(* IEC 61131-3 sources: daoli-st-library/DL_Process, 610 files *)

(* ---- FB_DL_AutoclaveSterilSeq.st ---- *)
(*==============================================================================
 * 组件名称 (Component)  : FB_DL_AutoclaveSterilSeq
 * 所属子库 (Sublibrary) : DL_Process
 * 当前版本 (Version)    : 1.0.1
 * 兼容性   (Platform)   : CODESYS 3.5+ / TwinCAT 3 / 汇川 InoProShop / 施耐德 Machine Expert
 *                         仅依赖 Standard.library（TON / R_TRIG / ABS），零厂商私有库
 * 功能描述 (Function)   : 灭菌釜脉动真空灭菌七态顺控（GMP F0 值合规）：
 *                           ePulse     脉动置换：重复「抽真空-进蒸汽」nPulseCnt 次
 *                                      （tPulse 半周期交替，回合完成计数）；
 *                           eHeatUp    升温：温压入带（fTempSetC±fTempTolC ∧
 *                                      fPrSetKpa±fPrTolKpa）→ eSteril，tHeatTo 超时
 *                                      分码 eNoPr（压不起）/ eNoTemp（温不到）；
 *                           eSteril    保压灭菌：tSteril 到时 ∧ F0 累计达标 ∧ 温压在带内
 *                                      才过相；F0 累计 fF0Acc += fF0Rate×fCycle/60，
 *                                      **带内才累加、带外冻结不倒扣**（保守侧）；
 *                                      带外持续 tBandTmo → eFault eSterilBand；
 *                           eExhaustDry 排气干燥 tExhaust 到时 → eDone。
 *                         bStop 任一相回 eIdle 不记故障；bStop 保留 F0 累计
 *                         （_fF0Acc 不清零，同批次再启动接续累计，仅 bReset
 *                         上升沿清 F0）；bReset 上升沿清全部锁存（R311）。
 * 接口     (Interface)  : 输入 bStart/bStop/bReset、fPrKpa 釜压（kPa）、fTempC 腔温（℃）、
 *                         fPrSetKpa/fTempSetC 灭菌设定、fPrTolKpa/fTempTolC 带半宽、
 *                         tSteril 保压时长、tPulse 脉动半周期、tHeatTo/tBandTmo/tExhaust
 *                         各相窗、nPulseCnt 置换次数、fF0Min F0 目标（min）、fF0Rate
 *                         F0 速率系数（min/min）、fCycle 扫描周期（s）；输出 ePhase 七态、
 *                         fF0AccMin F0 累计（min）、四相指示 BOOL 组、bDone、eCause、
 *                         bError。
 * 边界     (Boundary)   : ① **属主边界（写死）：本件只做灭菌时序编排与 F0 累计闸，不驱动
 *                         蒸汽阀/真空泵/排水阀**；执行器由 IO 映射层按相指示位驱动。
 *                         ② 七态 CASE + ELSE 兜底 eFault（R6）；段间 TON 各自专用
 *                         （tonPulse/tonHeatTo/tonSteril/tonBandTmo/tonExhaust，R228A
 *                         命名豁免式），段 0 无条件刷新，IN 由当前相与带内判据派生。
 *                         ③ eCause 分码：eNoPr（升不起压）/ eNoTemp（温不到）/ eSterilBand
 *                         （带外跌出）/ eCfgIllegal（组态非法）/ ePhaseBad（兜底），
 *                         归因唯一（R190）。
 *                         ④ 温压非有限 → eFault eCause=eNoTemp 分码（规格指定）。
 *                         ⑤ 组态闸：nPulseCnt=0、任一相时间 <= T#0S、设定值/带宽非正、
 *                         fF0Min<0、fF0Rate<0 → 锁存 eFault eCfgIllegal。
 *                         ⑥ F0 带外冻结：TON IN 派生式（带内才计时与累加），带外不倒扣
 *                         （头注释声明保守侧语义）。
 *                         ⑦ 温压带判定浮点全用 <= / >= 容差比较，禁 = 判等（R28）。
 *                         ⑧ 零全局耦合（无 GVL / VAR_EXTERNAL / 物理地址）。
 * 分工声明 (Scope)      : 温度带判定语义与 `FB_DL_ToleranceWindow` 同思想，本件自带实现
 *                         不引用（规格定为不内嵌引用，独立验收）。
 * 来源标签 (Source Tag) : T2-2 ◐（LBP 工艺分层只借灭菌工序分类事实，F0 累计口径为 GMP
 *                         公开定义，零文本复制）
 * 码表     (Codes)      : 本件不占用任何全局数字码位。出口为 ENUM 七态 + LREAL 累计 +
 *                         BOOL 组 + ENUM 成因；数字码位待主控收口阶段统一派号。
 * 红线自检 (Redline)    : R1 ✓ 零 GVL/VAR_EXTERNAL ｜ R2 ✓ 零 %I/%Q/%M ｜ R3 ✓ 纯 IEC 61131-3
 *                         R4 ✓ 非有限分码 + 带内累加闸 + 组态闸 + 周期缺省闸 ｜ R5 ✓ 声明逐行同行双语注释
 *                         R6 ✓ 七态 CASE 含 ELSE ｜ R7 ✓ 五 TON/两 R_TRIG 段 0 无条件刷新
 * 修订历史 (Revision)   : 2026-11-20  v1.0.1  R50 返修 R2：头注释补声明
 *                         「bStop 保留 F0 累计」口径——bStop 中止只清脉动
 *                         计数与子态，_fF0Acc 不清零（同批次再启动接续累计），
 *                         仅 bReset 上升沿清 F0 累计；逻辑零改动，契约不变。
 *                         2026-11-20  v1.0.0  R48 首版（批次 4 · 序号 18）
 *                         验收向量：脉动计满进升温；温压入带 + F0 达标 + tSteril 到 →
 *                         过相；带外跌出冻结计时；tBandTmo 超时故障；bStop 中止不记故障。
 *==============================================================================*)

TYPE E_DL_AcsPhase :
(
    eIdle      := 0,    // 待机 / Idle
    ePulse     := 10,   // 脉动置换相 / Pulsing vacuum-steam phase
    eHeatUp    := 20,   // 升温相 / Heat-up phase
    eSteril    := 30,   // 保压灭菌相 / Sterilization hold phase
    eExhaustDry:= 40,   // 排气干燥相 / Exhaust and dry phase
    eDone      := 50,   // 程序完成 / Sequence done
    eFault     := 90    // 故障（等复位）/ Fault, awaiting reset
);
END_TYPE

TYPE E_DL_AcsCause :
(
    eNone       := 0,   // 无异常 / No anomaly
    eNoPr       := 1,   // 升不起压（升温相压力超时）/ Pressure fail in heat-up
    eNoTemp     := 2,   // 温不到 / 温压非有限（分码共用温度侧成因）/ Temperature fail or non-finite
    eSterilBand := 3,   // 灭菌带外跌出超时 / Sterilization band dropout timeout
    eCfgIllegal := 4,   // 组态非法 / Illegal configuration
    ePhaseBad   := 5    // 非法相位兜底 / Illegal phase fallback
);
END_TYPE

FUNCTION_BLOCK FB_DL_AutoclaveSterilSeq
VAR_INPUT
    bStart    : BOOL := FALSE;     // 启动沿（eIdle 入脉动相） [-] / Start edge
    bStop     : BOOL := FALSE;     // 中止（任一相回 eIdle，不记故障） [-] / Abort to idle, no fault
    bReset    : BOOL := FALSE;     // 复位，上升沿清全部锁存（R311） [-] / Reset, rising edge clears all latches
    fPrKpa    : LREAL := 0.0;      // 釜压实测 [kPa] / Chamber pressure [kPa]
    fTempC    : LREAL := 0.0;      // 腔温实测 [℃] / Chamber temperature [degC]
    fPrSetKpa : LREAL := 200.0;    // 灭菌压力设定，域 > 0 [kPa] / Sterilization pressure setpoint [kPa]
    fTempSetC : LREAL := 121.0;    // 灭菌温度设定，域 > 0 [℃] / Sterilization temperature setpoint [degC]
    fPrTolKpa : LREAL := 10.0;     // 压力带半宽，域 > 0 [kPa] / Pressure band half-width [kPa]
    fTempTolC : LREAL := 1.0;      // 温度带半宽，域 > 0 [℃] / Temperature band half-width [degC]
    tSteril   : TIME := T#30M;     // 保压灭菌时长，域 > T#0S [ms] / Sterilization hold duration [ms]
    tPulse    : TIME := T#2M;      // 脉动半周期（抽真空/进蒸汽各一段），域 > T#0S [ms] / Pulse half-period [ms]
    tHeatTo   : TIME := T#60M;     // 升温相超时，域 > T#0S [ms] / Heat-up timeout [ms]
    tBandTmo  : TIME := T#5M;      // 灭菌带外容忍窗，域 > T#0S [ms] / Band dropout tolerance [ms]
    tExhaust  : TIME := T#15M;     // 排气干燥时长，域 > T#0S [ms] / Exhaust-dry duration [ms]
    nPulseCnt : UDINT := 3;        // 脉动置换次数，域 >= 1（=0 组态闸） [次] / Pulse swap count
    fF0Min    : LREAL := 3.0;      // F0 灭菌值目标，域 >= 0 [min] / F0 target [min]
    fF0Rate   : LREAL := 1.0;      // F0 累计速率系数（带内每分钟 F0 增量），域 >= 0 [min/min] / F0 rate coefficient
    fCycle    : LREAL := 0.0;      // 扫描周期（<=0 用缺省） [s] / Scan cycle, default used when <= 0
END_VAR
VAR_OUTPUT
    ePhase    : E_DL_AcsPhase;     // 当前相出口 [-] / Present phase outlet
    fF0AccMin : LREAL;             // F0 累计输出（带内累加、带外冻结） [min] / F0 accumulated [min]
    bPulseActive   : BOOL;         // 脉动相指示 [-] / Pulse phase indicator
    bHeatUpActive  : BOOL;         // 升温相指示 [-] / Heat-up phase indicator
    bSterilActive  : BOOL;         // 灭菌相指示 [-] / Sterilization phase indicator
    bExhaustActive : BOOL;         // 排气干燥相指示 [-] / Exhaust phase indicator
    bDone     : BOOL;              // 程序完成（eDone 驻留指示） [-] / Sequence done indicator
    eCause    : E_DL_AcsCause;     // 成因出口（锁存回放，R189） / Cause outlet, latched
    bError    : BOOL;              // 故障标志 [-] / Error flag
END_VAR
VAR
    _eState    : E_DL_AcsPhase := E_DL_AcsPhase.eIdle;   // 内部相（CASE 唯一写入目标） / Internal phase
    _eCause    : E_DL_AcsCause := E_DL_AcsCause.eNone;   // 成因锁存量 / Latched cause
    _bFault    : BOOL;             // 故障锁存位（解除沿 = bReset 上升沿） / Latched fault bit
    _nPulseDone: UDINT := 0;       // 脉动回合完成计数 [次] / Completed pulse swaps
    _bPulseStm : BOOL;             // 脉动子态（FALSE=抽真空段 / TRUE=进蒸汽段） / Pulse sub-state
    _bInBand   : BOOL;             // 当拍温压带内判据 [-] / In-band this scan
    _bNonFin   : BOOL;             // 温压非有限当拍量 [-] / Non-finite measurands this scan
    _bCfgBad   : BOOL;             // 组态非法当拍量 [-] / Illegal configuration this scan
    _fCy       : LREAL;            // 当拍有效周期 [s] / Effective cycle this scan
    _fF0Acc    : LREAL := 0.0;     // F0 累计锁存 [min] / F0 accumulator latch
    _bBusyPrev : BOOL;             // 上拍运行快照（bDone 迁出用） / Busy snapshot
    tonPulse   : TON;              // 脉动半周期定时器，段 0 无条件调用 / Pulse half-period timer
    tonHeatTo  : TON;              // 升温超时定时器，段 0 无条件调用 / Heat-up timeout timer
    tonSteril  : TON;              // 保压灭菌计时定时器，段 0 无条件调用 / Sterilization hold timer
    tonBandTmo : TON;              // 带外容忍窗定时器，段 0 无条件调用 / Band dropout tolerance timer
    tonExhaust : TON;              // 排气干燥计时定时器，段 0 无条件调用 / Exhaust-dry timer
    rtStart    : R_TRIG;           // 启动沿实例，段 0 无条件调用 / Start edge instance
    rtReset    : R_TRIG;           // 复位沿实例，段 0 无条件调用 / Reset edge instance
END_VAR
VAR CONSTANT
    DL_ACS_CYDEF : LREAL := 0.01;    // 缺省扫描周期 [s] / Default scan cycle
    DL_ACS_SEC   : LREAL := 60.0;    // 分秒换算基 [s/min] / Second-per-minute base
    DL_ACS_ZERO  : LREAL := 0.0;     // 非有限差值判零基准 [-] / Non-finite difference zero base
    DL_ACS_UDMAX : UDINT := 4294967295;   // UDINT 上限（脉动计数饱和点） [次] / UDINT ceiling
END_VAR

(* —— 段 0：非有限判 + 组态闸 + 周期派生 + 五 TON 两沿无条件周期刷新 —— *)
_bNonFin := (fPrKpa <> fPrKpa) OR ((fPrKpa - fPrKpa) <> DL_ACS_ZERO)
         OR (fTempC <> fTempC) OR ((fTempC - fTempC) <> DL_ACS_ZERO);   // 温压非有限（R245） / Non-finite pressure and temperature
_bCfgBad := (nPulseCnt = 0) OR (fPrSetKpa <= 0.0) OR (fTempSetC <= 0.0)
         OR (fPrTolKpa <= 0.0) OR (fTempTolC <= 0.0)
         OR (tSteril <= T#0S) OR (tPulse <= T#0S) OR (tHeatTo <= T#0S)
         OR (tBandTmo <= T#0S) OR (tExhaust <= T#0S)
         OR (fF0Min < 0.0) OR (fF0Rate < 0.0);          // 组态域闸（含 nPulseCnt=0） / Configuration gate
IF fCycle > 0.0 THEN
    _fCy := fCycle;                                     // 组态周期有效 / Configured cycle valid
ELSE
    _fCy := DL_ACS_CYDEF;                               // 周期缺省兜底 / Default cycle fallback
END_IF
rtStart(CLK := bStart);                                 // 启动沿，每拍必调 / Start edge, every scan
rtReset(CLK := bReset);                                 // 复位沿，每拍必调 / Reset edge, every scan
tonPulse(IN := (_eState = E_DL_AcsPhase.ePulse) AND (NOT tonPulse.Q), PT := tPulse);   // 脉动半周期自复位窗（R188） / Pulse self-reset window
tonHeatTo(IN := (_eState = E_DL_AcsPhase.eHeatUp), PT := tHeatTo);   // 升温超时（进相计时，出相自复位） / Heat-up timeout
tonSteril(IN := (_eState = E_DL_AcsPhase.eSteril) AND _bInBand, PT := tSteril);   // 灭菌计时（带内才计时，带外冻结） / Sterilization timer, in-band gated
tonBandTmo(IN := (_eState = E_DL_AcsPhase.eSteril) AND (NOT _bInBand), PT := tBandTmo);   // 带外容忍窗 / Band dropout tolerance
tonExhaust(IN := (_eState = E_DL_AcsPhase.eExhaustDry), PT := tExhaust);   // 排气干燥计时 / Exhaust timer

(* —— 段 1：带内判据（非有限按带外处理并分码 eNoTemp，先于 CASE 使用） —— *)
_bInBand := (NOT _bNonFin)
         AND (ABS(fTempC - fTempSetC) <= fTempTolC)     // 温度带内（容差比较，禁 =） / Temperature in band
         AND (ABS(fPrKpa - fPrSetKpa) <= fPrTolKpa);    // 压力带内 / Pressure in band

(* —— 段 2：单拍量预清零（_eState/_eCause/_bFault/_n PulseDone/_fF0Acc 锁存量不入清单，R107） —— *)
bPulseActive := FALSE;                                  // 脉动相指示预清 / Pulse indicator preset
bHeatUpActive := FALSE;                                 // 升温相指示预清 / Heat-up indicator preset
bSterilActive := FALSE;                                 // 灭菌相指示预清 / Sterilization indicator preset
bExhaustActive := FALSE;                                // 排气相指示预清 / Exhaust indicator preset
bDone := FALSE;                                         // 完成指示预清 / Done preset
bError := FALSE;                                        // 故障标志预清（R45 配对） / Error flag preset

(* —— 段 3：组态闸入故障 —— *)
IF _bCfgBad AND (NOT _bFault) THEN
    _bFault := TRUE;                                    // 锁存 / Latch
    _eCause := E_DL_AcsCause.eCfgIllegal;               // 归因：组态非法 / Cause: illegal config
    _eState := E_DL_AcsPhase.eFault;                    // 入故障相 / Enter fault
END_IF

(* —— 段 4：迁出链（bStop 优先不记故障；bReset 清全部锁存 R311） —— *)
IF bStop AND (_eState <> E_DL_AcsPhase.eIdle) THEN
    IF _eState = E_DL_AcsPhase.eFault THEN
        _bFault := FALSE;                               // 停机优先：故障相允许被停机清出 / Stop wins over fault
        _eCause := E_DL_AcsCause.eNone;                 // 清成因 / Clear cause
    END_IF
    _nPulseDone := 0;                                   // 清脉动计数 / Clear pulse count
    _bPulseStm := FALSE;                                // 清脉动子态 / Clear pulse sub-state
    _eState := E_DL_AcsPhase.eIdle;                     // 回待机（不记故障） / Back to idle, no fault
END_IF
IF rtReset.Q THEN
    _bFault := FALSE;                                   // 清故障锁存（R311） / Clear fault latch
    _eCause := E_DL_AcsCause.eNone;                     // 清成因 / Clear cause
    _nPulseDone := 0;                                   // 清脉动计数 / Clear pulse count
    _bPulseStm := FALSE;                                // 清脉动子态 / Clear pulse sub-state
    _fF0Acc := 0.0;                                     // 清 F0 累计 / Clear F0 accumulator
    _eState := E_DL_AcsPhase.eIdle;                     // 回待机 / Back to idle
END_IF

(* —— 段 5：七态顺控（只在无故障时推进；温压非有限 → 故障分码 eNoTemp） —— *)
IF (NOT _bFault) AND (NOT _bCfgBad) AND (NOT bStop) THEN
    IF _bNonFin AND (_eState <> E_DL_AcsPhase.eIdle) AND (_eState <> E_DL_AcsPhase.eDone) THEN
        _bFault := TRUE;                                // 运行相温压非有限：故障锁存（规格④） / Non-finite in running phase: fault
        _eCause := E_DL_AcsCause.eNoTemp;               // 归因分码：温度侧 / Cause: temperature side
        _eState := E_DL_AcsPhase.eFault;                // 入故障相 / Enter fault
    ELSE
        CASE _eState OF

        E_DL_AcsPhase.eIdle:
            IF rtStart.Q THEN
                _nPulseDone := 0;                       // 启动清脉动计数 / Clear pulse count on start
                _bPulseStm := FALSE;                    // 启动回抽真空子段 / Start in vacuum sub-phase
                _eState := E_DL_AcsPhase.ePulse;        // 入脉动相 / Enter pulse phase
            END_IF

        E_DL_AcsPhase.ePulse:
            IF tonPulse.Q THEN
                _bPulseStm := NOT _bPulseStm;           // 半周期到：抽真空/进蒸汽交替 / Half period: toggle sub-phase
                IF NOT _bPulseStm THEN
                    IF _nPulseDone < DL_ACS_UDMAX THEN
                        _nPulseDone := _nPulseDone + 1; // 完成一个完整回合（真空→蒸汽→真空）计数 / Count full swap round
                    END_IF
                END_IF
                IF _nPulseDone >= nPulseCnt THEN
                    _eState := E_DL_AcsPhase.eHeatUp;   // 置换次数达标：进升温相 / Swaps done: enter heat-up
                END_IF
            END_IF

        E_DL_AcsPhase.eHeatUp:
            IF _bInBand THEN
                _eState := E_DL_AcsPhase.eSteril;       // 温压入带：进保压灭菌相 / In band: enter sterilization
            ELSIF tonHeatTo.Q THEN
                IF ABS(fPrKpa - fPrSetKpa) > fPrTolKpa THEN
                    _eCause := E_DL_AcsCause.eNoPr;     // 压力超带：升不起压 / Pressure out of band: no pressure
                ELSE
                    _eCause := E_DL_AcsCause.eNoTemp;   // 压力入带而温度不达：温不到 / Temperature short
                END_IF
                _bFault := TRUE;                        // 超时故障锁存 / Latch fault
                _eState := E_DL_AcsPhase.eFault;        // 入故障相 / Enter fault
            END_IF

        E_DL_AcsPhase.eSteril:
            IF _bInBand THEN
                _fF0Acc := _fF0Acc + fF0Rate * _fCy / DL_ACS_SEC;   // 带内 F0 累计（速率×周期/60） / In-band F0 accumulation
            END_IF
            (* 带外不倒扣不累加（保守侧，头注释⑥）；带外容忍窗由 tonBandTmo 监视 *)
            IF tonBandTmo.Q THEN
                _eCause := E_DL_AcsCause.eSterilBand;   // 带外跌出超时 / Band dropout timeout
                _bFault := TRUE;                        // 锁存 / Latch
                _eState := E_DL_AcsPhase.eFault;        // 入故障相 / Enter fault
            ELSIF tonSteril.Q AND (_fF0Acc >= fF0Min) AND _bInBand THEN
                _eState := E_DL_AcsPhase.eExhaustDry;   // 计时到 ∧ F0 达标 ∧ 带内：过相（禁浮点 =，>= 判据） / Pass criteria met
            END_IF

        E_DL_AcsPhase.eExhaustDry:
            IF tonExhaust.Q THEN
                _eState := E_DL_AcsPhase.eDone;         // 排气干燥到时：进完成相 / Exhaust done: enter done
            END_IF

        E_DL_AcsPhase.eDone:
            ;                                           // 完成相驻留：由 bReset / bStop 迁出 / Held, exits via reset or stop

        E_DL_AcsPhase.eFault:
            ;                                           // 故障相驻留：由迁出链处理 / Held by exit chain

        ELSE
            _eCause := E_DL_AcsCause.ePhaseBad;         // 非法相位兜底归因 / Illegal phase cause
            _bFault := TRUE;                            // 锁存 / Latch
            _eState := E_DL_AcsPhase.eFault;            // 强拉故障相 / Force fault

        END_CASE
    END_IF
END_IF

(* —— 段 6：完成脉冲（由"运行→eDone"沿派生，单拍，R34 两段式） —— *)
IF _bBusyPrev AND (_eState = E_DL_AcsPhase.eDone) THEN
    bDone := TRUE;                                      // 程序完成单拍指示 / Done pulse
END_IF
_bBusyPrev := (_eState <> E_DL_AcsPhase.eIdle)
          AND (_eState <> E_DL_AcsPhase.eDone)
          AND (_eState <> E_DL_AcsPhase.eFault);        // 运行中快照（本拍末） / Busy snapshot at body end

(* —— 段 7：出口单点映射（相指示与相别同源，R191） —— *)
bPulseActive   := (_eState = E_DL_AcsPhase.ePulse);     // 脉动相指示 / Pulse indicator
bHeatUpActive  := (_eState = E_DL_AcsPhase.eHeatUp);    // 升温相指示 / Heat-up indicator
bSterilActive  := (_eState = E_DL_AcsPhase.eSteril);    // 灭菌相指示 / Sterilization indicator
bExhaustActive := (_eState = E_DL_AcsPhase.eExhaustDry);   // 排气相指示 / Exhaust indicator
IF _eState = E_DL_AcsPhase.eDone THEN
    bDone := TRUE;                                      // 完成相驻留期保持指示（R191 名实双出口声明） / Done held while resident
END_IF
ePhase := _eState;                                      // 当前相出口 / Present phase outlet
fF0AccMin := _fF0Acc;                                   // F0 累计出口 / F0 outlet
eCause := _eCause;                                      // 成因出口 / Cause outlet
bError := _bFault OR _bCfgBad;                          // 故障标志 = 锁存或组态非法 / Error = latch or config

END_FUNCTION_BLOCK

(* ---- FB_DL_BatchDoseSeq.st ---- *)
(*
    FB_DL_BatchDoseSeq —— 批次定量给料顺控（预给/快给/慢给/落料/校验 五相）
    ------------------------------------------------------------------
    组件名称  : FB_DL_BatchDoseSeq
    分类      : DL_Process / Batching
    前缀      : FB_DL_
    版本      : 1.0.0
    溯源      : 借鉴点 —— ISA-88（ANSI/ISA-88.00.01）批次控制模型的
                「单元配方 / 相逻辑 / 相超时 / 批次判定」分层思想，以及定量给料
                行业通行的三段给料法（快给料逼近 + 慢给料精给 + 落料补偿）。
                本件只借鉴**相划分与判定顺序**这两项公开语义。
                clean-room 声明 —— 零代码行复制；状态机为本件自有 ENUM + CASE，
                定时仅用 IEC 61131-3 标准库 TON，沿检测仅用标准库 R_TRIG。
                许可证 —— 本件 MIT；来源标签 isa88 指标准术语与模型，
                标准文本不属代码，无许可继承关系。
    平台      : 纯 IEC 61131-3，CODESYS 3.5 / TwinCAT 3 / InoProShop / Machine Expert 通用
    作者      : 道莅代码库 · PLC编程专家（R70 构建轮 · 批 1 · N4）
    ------------------------------------------------------------------
    功能说明  : 单批次定量给料顺控。相序：
                eIdle 待机 → ePreDose 预给料（预给料阀开，到 fPreW 止）
                → eFastDose 快给料（快给料阀开，到 fFastW 止）
                → eSlowDose 慢给料（慢给料阀开，到 fTarget - fFreeFall 止）
                → eSettle 落料（全阀关，等 tSettle 让空中料落下）
                → eCheck 校验（净重对 fTarget ± 公差带判定）
                → eComplete 完成（保持，等下一次 bStart）。
                超时归因唯一（R190）：预给 / 快给 / 慢给 / 落料四相各持独立码
                0303 / 0304 / 0305 / 0306，绝不共用同一枚举或同一码值。
                定时器设计：单实例 _tonPhase，PT 由当前相在段 4 以 IF/ELSIF 链
                逐相选择（含 ELSE 缺省），**每周期无条件调用**（规则 ⑦），
                故选相不依赖任何可能被跳过的分支；落料相的正常出口也复用该
                实例的 Q（PT = tSettle），故落料相不存在「正常完成」与「超时」
                两种语义，只有「到时间进入校验」一种。
                相内比较全部用 >= 的闭区间口径，不用浮点相等（规则 ④）。
    错误码    : 16#0002_0301 组态非法（阈值不单调 / 负公差 / 非有限），清锁存后回 eIdle —— 故障级
                16#0002_0302 称重值非有限，锁存并停料 —— 故障级
                16#0002_0303 预给料相超时 —— 故障级
                16#0002_0304 快给料相超时 —— 故障级
                16#0002_0305 慢给料相超时 —— 故障级
                16#0002_0306 落料相超时 —— 故障级
                16#0002_0307 欠重（净重低于 fTarget - fTolNeg）—— 故障级
                16#0002_0308 超重（净重高于 fTarget + fTolPos）—— 故障级
                16#0002_0309 非法相枚举值（CASE ELSE 兜底）—— 故障级
                16#0002_0310 启动被拒（称斗未回零，fWeight 超过 fZeroTol）—— 信息级，不置 bError
    码位总账  : 0301 / 0302 / 0303 / 0304 / 0305 / 0306 / 0307 / 0308 / 0309 用（均故障级）
                0310 用（信息级，bError 恒 FALSE）
    状态机    : ENUM E_DL_BdsPhase 八态，CASE 全覆盖 + ELSE 兜底（回 eFault 并置 0309）。
                迁移表见功能说明；bAbort 任意相 → eIdle（操作态，不发码）；
                bReset 上升沿：解锁存 → eIdle（仅此一条可到达的解除边，R188）。
    边界与披露: 一 组态判据逐项点名（R272）：fTarget / fPreW / fFastW / fFreeFall /
                   fTolNeg / fTolPos 全部纳入非有限闸，并校验单调链
                   0 < fPreW < fFastW < (fTarget - fFreeFall) 与 fFreeFall < fTarget、
                   两侧公差 >= 0；任一不满足即 0301 并锁存，**不落任何阈值比较**；
                二 称重输入非有限即锁存 0302，全部给料出口立即关断（失效安全方向）；
                三 失能语义：本件无 bEn 引脚，停机由 bAbort 承担 —— bAbort 为电平
                   有效，任意拍为 TRUE 即回 eIdle 且输出全清零，不发码（操作态）；
                四 出口语义（R191 名实双出口）：bUnder / bOver 为校验相判定结果位，
                   同时映射到故障码 0307 / 0308 并锁存；eComplete 为完成相标志，
                   完成不算故障，bError 恒 FALSE；
                五 bBusy 定义：给料 / 落料 / 校验三区间（真正占用设备的时间窗）；
                   bValid 定义：出口可信（未处在锁存故障相）；
                六 定时器 _tonPhase 与沿实例 _rtStart / _rtReset 均无条件周期调用；
                七 零全局变量、零 VAR_EXTERNAL、零物理地址、零数组下标、无除法。
    修订记录  : 2026-11-22 v1.0.0 首次入库（R70 构建轮 · 批 1 · N4）
*)
TYPE E_DL_BdsPhase :
(
    eIdle     := 0,   (* 待机，等待启动 / idle, waiting for a start *)
    ePreDose  := 10,  (* 预给料相（大流量阀开）/ the pre-dose phase, the coarse valve open *)
    eFastDose := 20,  (* 快给料相（快给料阀开）/ the fast-dose phase, the fast valve open *)
    eSlowDose := 30,  (* 慢给料相（慢给料阀开）/ the slow-dose phase, the fine valve open *)
    eSettle   := 40,  (* 落料相（全阀关，等空中料落下）/ the settling phase, all valves closed *)
    eCheck    := 50,  (* 校验相（净重对公差带判定）/ the check phase, the net weight against the tolerance *)
    eComplete := 60,  (* 完成相（保持到下次启动）/ the complete phase, held until the next start *)
    eFault    := 70   (* 故障相（锁存待复位）/ the fault phase, latched for a reset *)
);
END_TYPE

FUNCTION_BLOCK FB_DL_BatchDoseSeq
VAR_INPUT
    bStart    : BOOL := FALSE;             (* 启动命令（上升沿有效），[标志] / the start command, rising edge effective *)
    bAbort    : BOOL := FALSE;             (* 中止命令（电平有效），[标志] / the abort command, level effective *)
    bReset    : BOOL := FALSE;             (* 故障复位（上升沿有效），[标志] / the fault reset, rising edge effective *)
    fWeight   : LREAL := 0.0;              (* 称斗净重实时值，[kg] / the live net weight of the weigh hopper *)
    fTarget   : LREAL := 25.0;             (* 批次目标净重，[kg]，须 > 0 / the batch target weight, must be positive *)
    fPreW     : LREAL := 5.0;              (* 预给料结束重量点，[kg]，须 < fFastW / the pre-dose hand-over weight *)
    fFastW    : LREAL := 20.0;             (* 快给料结束重量点，[kg]，须 < fTarget - fFreeFall / the fast-dose hand-over weight *)
    fFreeFall : LREAL := 1.0;              (* 慢给料提前关断量（空中落差），[kg]，须 < fTarget / the in-flight cut-off weight *)
    fTolNeg   : LREAL := 0.2;              (* 允许负偏差，[kg]，须 >= 0 / the permitted negative deviation *)
    fTolPos   : LREAL := 0.2;              (* 允许正偏差，[kg]，须 >= 0 / the permitted positive deviation *)
    fZeroTol  : LREAL := 0.1;              (* 称斗空判定容差，[kg]，须 >= 0 / the empty-hopper tolerance *)
    tPre      : TIME := T#20S;             (* 预给料相超时，[ms] / the pre-dose phase timeout *)
    tFast     : TIME := T#30S;             (* 快给料相超时，[ms] / the fast-dose phase timeout *)
    tSlow     : TIME := T#30S;             (* 慢给料相超时，[ms] / the slow-dose phase timeout *)
    tSettle   : TIME := T#3S;              (* 落料稳定时间，[ms] / the settling duration *)
END_VAR
VAR_OUTPUT
    ePhase     : E_DL_BdsPhase := E_DL_BdsPhase.eIdle; (* 相状态出口，[相] / the phase outlet *)
    bPreOutlet : BOOL;                     (* 预给料阀 / 大流量出口命令，[标志] / the pre-dose outlet command *)
    bFastOutlet: BOOL;                     (* 快给料阀出口命令，[标志] / the fast-dose outlet command *)
    bSlowOutlet: BOOL;                     (* 慢给料阀出口命令，[标志] / the slow-dose outlet command *)
    bRunning   : BOOL;                     (* 批次进行中，[标志] / the batch is in progress *)
    bComplete  : BOOL;                     (* 批次完成（校验相通过后置位），[标志] / the batch completed *)
    bUnder     : BOOL;                     (* 欠重判定结果位，[标志] / the underweight verdict *)
    bOver      : BOOL;                     (* 超重判定结果位，[标志] / the overweight verdict *)
    fDeviation : LREAL;                    (* 实际偏差 fWeight - fTarget，[kg] / the actual deviation *)
    bBusy      : BOOL;                     (* 设备占用中（给料 / 落料 / 校验），[标志] / the equipment is occupied *)
    bValid     : BOOL;                     (* 出口可信（非锁存故障相），[标志] / the outlets are trustworthy *)
    bError     : BOOL;                     (* 故障标志，锁存故障时为 TRUE / the fault flag, raised while latched *)
    nErrCode   : UDINT;                    (* 错误码，0 = 正常，锁存回放 / the error id, 0 = ok, replayed from the latch *)
END_VAR
VAR
    _rtStart     : R_TRIG;                 (* 启动上升沿实例（无条件调用）/ the start rising edge instance *)
    _rtReset     : R_TRIG;                 (* 复位上升沿实例（无条件调用）/ the reset rising edge instance *)
    _tonPhase    : TON;                    (* 相计时 / 落料计时实例（无条件调用）/ the phase and settle timer *)
    _ePhase      : E_DL_BdsPhase := E_DL_BdsPhase.eIdle; (* 相状态寄存器，[相] / the internal phase register *)
    _bFault      : BOOL;                   (* 故障锁存位，仅 bReset 上升沿解除 / the latched fault bit *)
    _nCodeLatch  : UDINT;                  (* 锁存成因码，故障期回放 / the latched cause code, replayed *)
    _bCfgBad     : BOOL;                   (* 组态非法标志（逐拍重算）/ the configuration fault flag *)
    _bInBad      : BOOL;                   (* 称重非有限标志（逐拍重算）/ the weight fault flag *)
    _bTimerIn    : BOOL;                   (* 相计时器 IN 条件（显式条件，段 4 计算）/ the timer IN condition *)
    _tPhasePt    : TIME;                   (* 相计时器 PT 当前值（逐相选择）/ the timer PT for the current phase *)
    _bStartOk    : BOOL;                   (* 启动前置条件成立（称斗已空）/ the start precondition holds *)
    _fSlowCut    : LREAL;                  (* 慢给料关断重量点 = fTarget - fFreeFall，[kg] / the slow-dose cut-off weight *)
    _fDev        : LREAL;                  (* 偏差中间量，[kg] / the deviation temporary *)
END_VAR
VAR CONSTANT
    DL_BDS_FMAX  : LREAL := 1.0E30;        (* 非有限筛查幅值上限，[kg] / the finiteness screening cap *)
    DL_BDS_UNDER : UDINT := 16#0002_0307;  (* 欠重码字面量（CASE 内引用，避免魔数）/ the underweight literal *)
    DL_BDS_OVER  : UDINT := 16#0002_0308;  (* 超重码字面量 / the overweight literal *)
END_VAR

// 段 1｜出口预置（R256 统一出口预置 + 单拍位两段式的第一段）/ segment 1, preset every outlet
ePhase      := _ePhase;                    // 相出口先镜像寄存器 / mirror the phase register first
bPreOutlet  := FALSE;                      // 预给料出口预清零 / preset the pre-dose outlet false
bFastOutlet := FALSE;                      // 快给料出口预清零 / preset the fast-dose outlet false
bSlowOutlet := FALSE;                      // 慢给料出口预清零 / preset the slow-dose outlet false
bRunning    := FALSE;                      // 运行标志预清零 / preset the running flag false
bComplete   := FALSE;                      // 完成标志预清零 / preset the complete flag false
bUnder      := FALSE;                      // 欠重结果预清零 / preset the underweight verdict false
bOver       := FALSE;                      // 超重结果预清零 / preset the overweight verdict false
fDeviation  := 0.0;                        // 偏差预置零 / preset the deviation to zero
bBusy       := FALSE;                      // 占用标志预清零 / preset the busy flag false
bValid      := TRUE;                       // 可用标志预置真（故障相再清）/ preset valid true, cleared in the fault phase
bError      := FALSE;                      // 故障标志预清零 / preset the error flag false
nErrCode    := 0;                          // 错误码预置无错 / preset the code to zero
_bTimerIn   := FALSE;                      // 计时条件预清零 / preset the timer condition false
_tPhasePt   := tPre;                       // 计时 PT 预置缺省值 / preset the timer PT to the default

// 段 2｜沿检测实例无条件调用（规则 ⑦）/ segment 2, the edge instances, called unconditionally
_rtStart(CLK := bStart);                   // 启动沿，每周期无条件刷新 / the start edge, refreshed every scan
_rtReset(CLK := bReset);                   // 复位沿，每周期无条件刷新 / the reset edge, refreshed every scan

// 段 3｜复位解除：唯一可到达的锁存解除边（R188）/ segment 3, the only latch release edge
IF _rtReset.Q THEN                         // 复位上升沿 / the reset rising edge
    _bFault     := FALSE;                  // 解除故障锁存 / release the fault latch
    _nCodeLatch := 0;                      // 清锁存码 / clear the latched code
    _ePhase     := E_DL_BdsPhase.eIdle;    // 回待机相（安全相）/ back to the safe idle phase
END_IF

// 段 4｜组态守卫（阈值单调链 + 公差非负 + 全量非有限闸，R272）/ segment 4, the configuration guard
_fSlowCut := fTarget - fFreeFall;          // 慢给料关断点，供单调链复检 / the slow-dose cut-off point
_bCfgBad := (fTarget <= 0.0)                                             // 目标非正 / a non positive target
         OR (fFreeFall < 0.0)                                            // 落差为负 / a negative in-flight weight
         OR (fFreeFall >= fTarget)                                       // 落差吞没目标 / the in-flight swallows the target
         OR (fPreW <= 0.0)                                               // 预给料点非正 / a non positive pre-dose point
         OR (fFastW <= fPreW)                                            // 快给料点未高于预给料点 / the fast point not above the pre point
         OR (fFastW >= _fSlowCut)                                        // 快给料点越过慢给料关断点 / the fast point over the slow cut-off
         OR (fTolNeg < 0.0)                                              // 负公差为负 / a negative tolerance
         OR (fTolPos < 0.0)                                              // 正公差为负 / a negative tolerance
         OR (fZeroTol < 0.0)                                             // 空斗容差为负 / a negative empty tolerance
         OR (fTarget <> fTarget) OR ((fTarget - fTarget) <> 0.0) OR (ABS(fTarget) > DL_BDS_FMAX)
         OR (fPreW <> fPreW) OR ((fPreW - fPreW) <> 0.0) OR (ABS(fPreW) > DL_BDS_FMAX)
         OR (fFastW <> fFastW) OR ((fFastW - fFastW) <> 0.0) OR (ABS(fFastW) > DL_BDS_FMAX)
         OR (fFreeFall <> fFreeFall) OR ((fFreeFall - fFreeFall) <> 0.0) OR (ABS(fFreeFall) > DL_BDS_FMAX)
         OR (fTolNeg <> fTolNeg) OR ((fTolNeg - fTolNeg) <> 0.0) OR (ABS(fTolNeg) > DL_BDS_FMAX)
         OR (fTolPos <> fTolPos) OR ((fTolPos - fTolPos) <> 0.0) OR (ABS(fTolPos) > DL_BDS_FMAX)
         OR (fZeroTol <> fZeroTol) OR ((fZeroTol - fZeroTol) <> 0.0) OR (ABS(fZeroTol) > DL_BDS_FMAX);

// 段 5｜输入守卫：称重非有限 / segment 5, the weight input guard
_bInBad := (fWeight <> fWeight) OR ((fWeight - fWeight) <> 0.0) OR (ABS(fWeight) > DL_BDS_FMAX);

// 段 6｜首次成因锁存（故障期不重推断，回放锁存码，R189）/ segment 6, the first-cause latch
IF NOT _bFault THEN                        // 未锁存才登记成因 / a cause is registered only while not latched
    IF _bCfgBad THEN                       // 组态非法优先归因（根因）/ the configuration first, it is the root cause
        _bFault     := TRUE;               // 置锁存 / latch it
        _nCodeLatch := 16#0002_0301;       // 故障级：组态非法 / fault level: an illegal configuration
        _ePhase     := E_DL_BdsPhase.eFault; // 迁入故障相 / enter the fault phase
    ELSIF _bInBad THEN                     // 称重非有限 / the weight is non finite
        _bFault     := TRUE;               // 置锁存 / latch it
        _nCodeLatch := 16#0002_0302;       // 故障级：输入非有限 / fault level: the input is non finite
        _ePhase     := E_DL_BdsPhase.eFault; // 迁入故障相 / enter the fault phase
    END_IF
END_IF

// 段 7｜中止命令（操作态，不发码）：任意相回待机 / segment 7, the abort command, an operator state
IF bAbort AND NOT _bFault THEN             // 中止有效且无锁存故障 / an abort without a latched fault
    _ePhase := E_DL_BdsPhase.eIdle;        // 回待机（安全相）/ back to the safe idle phase
END_IF

// 段 8｜相计时器 PT 选择与无条件调用（规则 ⑦，选相不依赖可跳过分支）/ segment 8, the timer PT selection and the unconditional call
IF _ePhase = E_DL_BdsPhase.ePreDose THEN       // 预给料相 / the pre-dose phase
    _tPhasePt := tPre;                         // 预给料超时值 / the pre-dose timeout
    _bTimerIn := TRUE;                         // 相内计时有效 / the timer runs inside the phase
ELSIF _ePhase = E_DL_BdsPhase.eFastDose THEN   // 快给料相 / the fast-dose phase
    _tPhasePt := tFast;                        // 快给料超时值 / the fast-dose timeout
    _bTimerIn := TRUE;                         // 相内计时有效 / the timer runs
ELSIF _ePhase = E_DL_BdsPhase.eSlowDose THEN   // 慢给料相 / the slow-dose phase
    _tPhasePt := tSlow;                        // 慢给料超时值 / the slow-dose timeout
    _bTimerIn := TRUE;                         // 相内计时有效 / the timer runs
ELSIF _ePhase = E_DL_BdsPhase.eSettle THEN     // 落料相 / the settling phase
    _tPhasePt := tSettle;                      // 落料时长即其正常出口 / the settling duration is its normal exit
    _bTimerIn := TRUE;                         // 落料计时有效 / the timer runs
ELSE                                           // 其余相不参与计时（缺省分支，非状态机的 ELSE）/ the other phases do not time
    _tPhasePt := tPre;                         // 缺省 PT，保证 PT 恒有定义 / a default PT, always defined
    _bTimerIn := FALSE;                        // 计时条件清零 / the timer condition cleared
END_IF
_tonPhase(IN := _bTimerIn, PT := _tPhasePt);   // 每周期无条件调用 / called every scan without exception

// 段 9｜相状态机（ENUM + CASE + ELSE 兜底）/ segment 9, the phase machine
CASE _ePhase OF
    E_DL_BdsPhase.eIdle:                        // 待机相 / the idle phase
        bValid := TRUE;                         // 待机出口可信 / the idle outlets are trustworthy
        IF _rtStart.Q AND NOT _bFault THEN      // 启动沿且无锁存故障 / a start edge without a latched fault
            _bStartOk := (fWeight <= fZeroTol); // 前置条件：称斗已空 / the precondition, an empty hopper
            IF _bStartOk THEN                   // 前置成立 / the precondition holds
                _ePhase := E_DL_BdsPhase.ePreDose; // 进入预给料相 / enter the pre-dose phase
            ELSE                                // 称斗有残料 / the hopper is not empty
                nErrCode := 16#0002_0310;       // 信息级：启动被拒（不置 bError，R45）/ info level: the start is refused
                _ePhase  := E_DL_BdsPhase.eIdle; // 保持待机 / stay idle
            END_IF
        END_IF
    E_DL_BdsPhase.ePreDose:                     // 预给料相 / the pre-dose phase
        bRunning   := TRUE;                     // 批次进行中 / the batch runs
        bBusy      := TRUE;                     // 设备占用 / the equipment is occupied
        bPreOutlet := TRUE;                     // 预给料阀开 / open the pre-dose outlet
        IF fWeight >= fPreW THEN                // 到达预给料结束重量 / the pre-dose hand-over weight reached
            _ePhase := E_DL_BdsPhase.eFastDose; // 进入快给料相 / enter the fast-dose phase
        ELSIF _tonPhase.Q THEN                  // 相超时（归因唯一 0303）/ the phase timed out
            _bFault     := TRUE;                // 锁存故障 / latch the fault
            _nCodeLatch := 16#0002_0303;        // 故障级：预给料超时 / fault level: the pre-dose timed out
            _ePhase     := E_DL_BdsPhase.eFault; // 迁入故障相 / enter the fault phase
        END_IF
    E_DL_BdsPhase.eFastDose:                    // 快给料相 / the fast-dose phase
        bRunning    := TRUE;                    // 批次进行中 / the batch runs
        bBusy       := TRUE;                    // 设备占用 / occupied
        bFastOutlet := TRUE;                    // 快给料阀开 / open the fast-dose outlet
        IF fWeight >= fFastW THEN               // 到达快给料结束重量 / the fast-dose hand-over weight reached
            _ePhase := E_DL_BdsPhase.eSlowDose; // 进入慢给料相 / enter the slow-dose phase
        ELSIF _tonPhase.Q THEN                  // 相超时（归因唯一 0304）/ the phase timed out
            _bFault     := TRUE;                // 锁存故障 / latch the fault
            _nCodeLatch := 16#0002_0304;        // 故障级：快给料超时 / fault level: the fast-dose timed out
            _ePhase     := E_DL_BdsPhase.eFault; // 迁入故障相 / enter the fault phase
        END_IF
    E_DL_BdsPhase.eSlowDose:                    // 慢给料相 / the slow-dose phase
        bRunning    := TRUE;                    // 批次进行中 / the batch runs
        bBusy       := TRUE;                    // 设备占用 / occupied
        bSlowOutlet := TRUE;                    // 慢给料阀开 / open the slow-dose outlet
        IF fWeight >= _fSlowCut THEN            // 到达提前关断点（含空落差补偿）/ the cut-off point reached
            _ePhase := E_DL_BdsPhase.eSettle;   // 进入落料相 / enter the settling phase
        ELSIF _tonPhase.Q THEN                  // 相超时（归因唯一 0305）/ the phase timed out
            _bFault     := TRUE;                // 锁存故障 / latch the fault
            _nCodeLatch := 16#0002_0305;        // 故障级：慢给料超时 / fault level: the slow-dose timed out
            _ePhase     := E_DL_BdsPhase.eFault; // 迁入故障相 / enter the fault phase
        END_IF
    E_DL_BdsPhase.eSettle:                      // 落料相（全阀关）/ the settling phase, all outlets closed
        bRunning := TRUE;                       // 批次进行中 / the batch runs
        bBusy    := TRUE;                       // 设备占用 / occupied
        IF _tonPhase.Q THEN                     // 落料时长到（正常出口，非超时）/ the settling done, the normal exit
            _ePhase := E_DL_BdsPhase.eCheck;    // 进入校验相 / enter the check phase
        END_IF
    E_DL_BdsPhase.eCheck:                       // 校验相 / the check phase
        bRunning   := TRUE;                     // 批次进行中 / the batch runs
        bBusy      := TRUE;                     // 设备占用 / occupied
        _fDev      := fWeight - fTarget;        // 实际偏差 / the actual deviation
        fDeviation := _fDev;                    // 偏差出口 / the deviation outlet
        IF _fDev < (0.0 - fTolNeg) THEN         // 欠重（低于负公差）/ underweight
            bUnder      := TRUE;                // 欠重结果位 / the underweight verdict
            _bFault     := TRUE;                // 锁存故障 / latch the fault
            _nCodeLatch := DL_BDS_UNDER;        // 故障级：欠重 / fault level: underweight
            _ePhase     := E_DL_BdsPhase.eFault; // 迁入故障相 / enter the fault phase
        ELSIF _fDev > fTolPos THEN              // 超重（高于正公差）/ overweight
            bOver       := TRUE;                // 超重结果位 / the overweight verdict
            _bFault     := TRUE;                // 锁存故障 / latch the fault
            _nCodeLatch := DL_BDS_OVER;         // 故障级：超重 / fault level: overweight
            _ePhase     := E_DL_BdsPhase.eFault; // 迁入故障相 / enter the fault phase
        ELSE                                    // 落在公差带内 / inside the tolerance band
            _ePhase := E_DL_BdsPhase.eComplete; // 进入完成相 / enter the complete phase
        END_IF
    E_DL_BdsPhase.eComplete:                    // 完成相（保持）/ the complete phase, held
        bComplete := TRUE;                      // 完成标志 / the complete flag
        bValid    := TRUE;                      // 完成相出口可信 / the complete outlets are trustworthy
        IF _rtStart.Q AND (fWeight <= fZeroTol) THEN // 称斗已卸空且再次启动 / the hopper emptied and a start arrived
            _ePhase := E_DL_BdsPhase.ePreDose;  // 直接进入下一批预给料 / start the next batch
        END_IF
    E_DL_BdsPhase.eFault:                       // 故障相（锁存保持）/ the fault phase, latched
        bValid   := FALSE;                      // 出口不可信 / the outlets are not trustworthy
        bError   := TRUE;                       // 故障标志置位 / raise the fault flag
        nErrCode := _nCodeLatch;                // 回放锁存码（不按当下输入重推断）/ replay the latched code
    ELSE                                        // 非法枚举兜底（回安全相 + 置码，规则 ⑥）/ the illegal enumeration guard
        _bFault     := TRUE;                    // 置锁存 / latch it
        _nCodeLatch := 16#0002_0309;            // 故障级：非法相枚举 / fault level: an illegal phase value
        _ePhase     := E_DL_BdsPhase.eFault;    // 回安全相（故障相）/ force the safe fault phase
        bValid      := FALSE;                   // 出口不可信 / the outlets are not trustworthy
        bError      := TRUE;                    // 故障标志置位（禁静默）/ raise the fault flag
        nErrCode    := _nCodeLatch;             // 回放锁存码 / replay the latched code
END_CASE

// 段 10｜相出口映射（名实双出口同源，R191）/ segment 10, the phase outlet mapping
ePhase := _ePhase;                          // 相出口 = 寄存器（单点写入，段 9 之后不再触碰）/ the phase outlet mirrors the register
END_FUNCTION_BLOCK

(* ---- FB_DL_ChamberPumpDownSeq.st ---- *)
(*==============================================================================
 * 组件名称 (Component)  : FB_DL_ChamberPumpDownSeq
 * 所属子库 (Sublibrary) : DL_Process
 * 当前版本 (Version)    : 1.0.0
 * 兼容性   (Platform)   : CODESYS 3.5+ / TwinCAT 3 / 汇川 InoProShop / 施耐德 Machine Expert
 *                         仅依赖 Standard.library（TON / R_TRIG），零厂商私有库
 * 功能描述 (Function)   : 腔体抽真空顺控与漏率复测（四段：抽气 → 稳压 → 漏率复测 → 放气限速）。
 *                         每相一枚**专用** TON，PT 各绑一个时间引脚，绝不复用实例改 PT：
 *                           ePump   抽气  ：tonPumpTo  PT = tPumpTo  （到目标真空 fPrTargetKpa 即过相）
 *                           eStab   稳压  ：tonStabTo  PT = tStab    （纯定时过相）
 *                           eLeak   复测  ：tonLeakWin PT = tLeakWin （窗满即算漏率）
 *                           eVent   放气  ：tonVentTo  PT = tVentTo  （到常压即回待机）
 *                         **漏率判据**：窗起压 fPrStart 与窗末压 fPrEnd 之差除以窗内实际时长；
 *                         窗内实际时长＝采样计数 × 采样周期（fSampleS），因此不需要 TIME→实数转换
 *                         （规避跨平台时间转换链，R64 家族），且分母双闸（计数 ≥ 1 且周期 > 0）。
 *                         **放气限速**：逐拍放气速率超 fVentRateMaxKpaPerS 时当拍关阀（bang-bang 限速），
 *                         并在下一拍重新开阀，形成占空比式限速；超速不锁存（工艺可容忍），只置信息级。
 *                         验收向量：
 *                           ① 目标 −90 kPa，实测 −90.2 → 过相进入稳压
 *                           ② 窗 5 s、周期 0.1 s、Δp = 0.5 kPa → 漏率 0.5/(50×0.1) = 0.1 kPa/s
 *                           ③ fLeakMax = 0.05 kPa/s 且实测 0.1 → eLeakNg 锁存，禁止进入放气
 *                           ④ 放气速率 2.0 kPa/s > 上限 1.0 → 当拍关阀 + eVentTooFast（信息级）
 * 接口     (Interface)  : 入 bStart 启动沿、fPrMeasKpa 实测腔压、fPrTargetKpa 目标真空（负值）、
 *                         fLeakMaxKpaPerS 漏率上限、fVentRateMaxKpaPerS 放气速率上限、fSampleS 采样周期、
 *                         tPumpTo / tStab / tLeakWin / tVentTo 四段时间、bStop 中止、bReset 复位沿；
 *                         出 bPumpValve 抽气阀位、bVentValve 放气阀位、fLeakRateKpaPerS 实测漏率、
 *                         bLeakNg 漏率超限锁存、bBusy 顺控中、bDone 完成脉冲（单拍）、
 *                         ePhase 当前相、eCause 成因、bError 故障标志。
 * 边界     (Boundary)   : ① **属主边界（写死）：本件只做"腔体抽真空时序 + 漏率判据 + 放气限速"，
 *                         不驱动真空泵/角阀线圈、不做脱泡/灌胶工艺**——灌胶真空脱泡四相属
 *                         `FB_DL_ModulePottingVac`，两件不同属主、判据不共用（R47 边界声明）；
 *                         ② **分母双闸**：窗内采样计数 = 0 或采样周期 ≤ 0 时漏率判据整段不判，
 *                         并锁存 eCfgIllegal（静默失效比报错危险，R179）；
 *                         ③ **组态闸**：四段时间须 > T#0S、目标真空须 < 0（相对压）、
 *                         两上限须 > 0，违反即锁存 eCfgIllegal；
 *                         ④ **一相一 TON**：四枚专用 TON 段 0 无条件调用，IN 由当前相派生
 *                         （R228A/R275），无跨相累积；
 *                         ⑤ **eFault 可迁出**：bReset 上升沿 → eIdle；bStop 在非故障相回 eIdle
 *                         并置中止脉冲（泵/阀在出口侧随相切断）；
 *                         ⑥ 零全局耦合、零物理地址。
 * 分工声明 (Scope)      : 本件只管"腔体抽真空与漏率复测"。不接管：灌胶脱泡四相
 *                         （属 FB_DL_ModulePottingVac）、真空泵轮换（属泵组件）、
 *                         腔体压力闭环调节（属压力环件）。
 * 来源标签 (Source Tag) : ROADMAP 空勾真缺口 P1（腔体抽真空与漏率复测，自研 clean-room）
 * 码表     (Codes)      : 本件不占用任何全局数字码位（零码位范式 R297）；诊断由 BOOL + ENUM 出口承担。
 * 红线自检 (Redline)    : R1 ✓ 零 GVL/VAR_EXTERNAL ｜ R2 ✓ 零 %I/%Q/%M ｜ R3 ✓ 纯 IEC 61131-3
 *                         R4 ✓ 分母双闸 + 组态闸 + 漏率钳位 + 非有限闸 ｜ R5 ✓ 声明逐行同行双语注释
 *                         R6 ✓ ENUM+CASE 含 ELSE 兜底 ｜ R7 ✓ 四 TON/两 R_TRIG 段 0 无条件刷新
 * 修订历史 (Revision)   : 2026-11-19  v1.0.0  R47 首版（批次 3 · 序号 14）
 *==============================================================================*)

TYPE E_DL_CpdPhase :
(
    eIdle  := 0,    // 待机相（泵/阀全停） / Idle, pump and valves off
    ePump  := 10,   // 抽气相（等到目标真空） / Pumping down to the target
    eStab  := 20,   // 稳压相（压力稳定） / Stabilising
    eLeak  := 30,   // 漏率复测相（测量窗内） / Leak-rate measurement window
    eVent  := 40,   // 放气相（限速） / Venting with rate limiting
    eFault := 90    // 故障相（等复位） / Fault, awaiting reset
);
END_TYPE

TYPE E_DL_CpdCause :
(
    eNone         := 0,   // 无异常 / No anomaly
    eCfgIllegal   := 1,   // 组态非法（时间/目标/上限/采样越域） / Illegal configuration
    ePumpTimeout  := 2,   // 抽气超时未达目标真空 / Pump-down timeout
    eLeakNg       := 3,   // 漏率超限（锁存） / Leak rate exceeded, latched
    eVentTimeout  := 4,   // 放气超时未到常压 / Vent timeout
    eVentTooFast  := 5,   // 放气速率超限（信息级，当拍关阀） / Vent rate exceeded, info level
    ePhaseBad     := 6    // 非法相位兜底 / Illegal phase fallback
);
END_TYPE

FUNCTION_BLOCK FB_DL_ChamberPumpDownSeq
VAR_INPUT
    bStart             : BOOL := FALSE;     // 启动沿，进入抽气相 [-] / Start edge, enters pumping
    bStop              : BOOL := FALSE;     // 中止（非故障相回待机） [-] / Abort
    fPrMeasKpa         : LREAL := 0.0;      // 实测腔压（相对压，负值为真空） [kPa] / Measured chamber pressure [kPa]
    fPrTargetKpa       : LREAL := -90.0;    // 目标真空，域 < 0 [kPa] / Target vacuum, < 0
    fLeakMaxKpaPerS    : LREAL := 0.05;     // 漏率上限，域 > 0 [kPa/s] / Leak-rate limit, > 0
    fVentRateMaxKpaPerS: LREAL := 1.0;      // 放气速率上限，域 > 0 [kPa/s] / Vent-rate limit, > 0
    fSampleS           : LREAL := 0.1;      // 调用采样周期，域 > 0 [s] / Sampling period, > 0
    tPumpTo            : TIME := T#120S;    // 抽气超时，域 > T#0S [ms] / Pump-down timeout
    tStab              : TIME := T#5S;      // 稳压时长，域 > T#0S [ms] / Stabilisation time
    tLeakWin           : TIME := T#10S;     // 漏率测量窗，域 > T#0S [ms] / Leak measurement window
    tVentTo            : TIME := T#60S;     // 放气超时，域 > T#0S [ms] / Vent timeout
    bReset             : BOOL := FALSE;     // 故障复位沿 [-] / Fault reset edge
END_VAR
VAR_OUTPUT
    bPumpValve  : BOOL := FALSE;                          // 抽气阀位（含真空泵启动允许） [-] / Pump valve position
    bVentValve  : BOOL := FALSE;                          // 放气阀位 [-] / Vent valve position
    fLeakRateKpaPerS : LREAL := 0.0;                      // 实测漏率 [kPa/s] / Measured leak rate [kPa/s]
    bLeakNg     : BOOL := FALSE;                          // 漏率超限锁存（等复位） [-] / Leak NG, latched
    bBusy       : BOOL := FALSE;                          // 顺控进行中 [-] / Sequence busy
    bDone       : BOOL := FALSE;                          // 完成脉冲（单拍） [-] / Completion pulse, single scan
    bAborted    : BOOL := FALSE;                          // 中止脉冲（单拍） [-] / Abort pulse, single scan
    ePhase      : E_DL_CpdPhase := E_DL_CpdPhase.eIdle;   // 当前相出口 [-] / Present phase outlet
    eCause      : E_DL_CpdCause := E_DL_CpdCause.eNone;   // 成因出口（R190 归因唯一） [-] / Cause outlet
    bError      : BOOL := FALSE;                          // 故障标志（仅故障级成因） [-] / Error flag, fault level only
END_VAR
VAR
    _eState    : E_DL_CpdPhase := E_DL_CpdPhase.eIdle;    // 内部相（CASE 唯一写入目标） / Internal phase
    _eCause    : E_DL_CpdCause := E_DL_CpdCause.eNone;    // 成因锁存量 / Latched cause
    _bFault    : BOOL := FALSE;                           // 故障锁存位 / Latched fault bit
    _bLeakNg   : BOOL := FALSE;                           // 漏率超限锁存位 / Latched leak-NG bit
    _bDone     : BOOL := FALSE;                           // 完成脉冲内部位（单拍） / Internal completion pulse
    _bAborted  : BOOL := FALSE;                           // 中止脉冲内部位（单拍） / Internal abort pulse
    _bBusyPrev : BOOL := FALSE;                           // 上拍忙碌快照 / Busy snapshot of the previous scan
    _fPrStart  : LREAL := 0.0;                            // 测量窗起始压力 [kPa] / Pressure at the window start
    _fPrPrev   : LREAL := 0.0;                            // 上拍压力（放气速率用） [kPa] / Previous pressure for the vent rate
    _fPrNow    : LREAL := 0.0;                            // 当拍压力工作值 [kPa] / Pressure working value
    _fRate     : LREAL := 0.0;                            // 速率工作值 [kPa/s] / Rate working value
    _fDtS      : LREAL := 0.0;                            // 实际时长（计数 × 周期） [s] / Effective duration [s]
    _nWinCnt   : UDINT := 0;                              // 窗内采样计数 [个] / Sample count inside the window
    _bCfgBad   : BOOL := FALSE;                           // 组态非法当拍量 / Illegal configuration this scan
    _bPrOk     : BOOL := FALSE;                           // 压力样本有限性结论 / Pressure sample finiteness
    _bVent     : BOOL := FALSE;                           // 放气阀内部位（限速判决，单拍重算） / Internal vent valve bit
    tonPumpTo  : TON;                                     // 抽气相专用超时，段 0 无条件调用 / Pump dedicated timeout
    tonStabTo  : TON;                                     // 稳压相专用时长，段 0 无条件调用 / Stabilisation dedicated time
    tonLeakWin : TON;                                     // 复测相专用窗，段 0 无条件调用 / Leak-window dedicated timer
    tonVentTo  : TON;                                     // 放气相专用超时，段 0 无条件调用 / Vent dedicated timeout
    rtStart    : R_TRIG;                                  // 启动沿实例，段 0 无条件调用 / Start edge instance
    rtReset    : R_TRIG;                                  // 复位沿实例，段 0 无条件调用 / Reset edge instance
END_VAR
VAR CONSTANT
    DL_CPD_EPS : LREAL := 1.0E-9;         // 浮点判等容差 [kPa] / Equality tolerance [kPa]
END_VAR

(* —— 段 0：组态闸 + 四枚专用 TON 与两沿无条件周期刷新（R228A/R275） —— *)
_bCfgBad := (tPumpTo <= T#0S) OR (tStab <= T#0S) OR (tLeakWin <= T#0S) OR (tVentTo <= T#0S)   // 四时间须为正 / Four times positive
         OR (fPrTargetKpa >= 0.0)                                                              // 目标真空须为负（相对压） / Target vacuum negative
         OR (fLeakMaxKpaPerS <= 0.0) OR (fVentRateMaxKpaPerS <= 0.0)                           // 两上限须为正 / Both limits positive
         OR (fSampleS <= 0.0) OR (fSampleS <> fSampleS);                                        // 采样周期须为正且有限 / Sampling period positive and finite
rtStart(CLK := bStart);                                                                        // 启动沿 / Start edge
rtReset(CLK := bReset);                                                                        // 复位沿 / Reset edge
tonPumpTo(IN := (_eState = E_DL_CpdPhase.ePump), PT := tPumpTo);                                // 抽气相专用超时 / Pump timeout
tonStabTo(IN := (_eState = E_DL_CpdPhase.eStab), PT := tStab);                                  // 稳压相专用时长 / Stabilisation time
tonLeakWin(IN := (_eState = E_DL_CpdPhase.eLeak), PT := tLeakWin);                              // 复测相专用窗 / Leak window
tonVentTo(IN := (_eState = E_DL_CpdPhase.eVent), PT := tVentTo);                                // 放气相专用超时 / Vent timeout

(* —— 段 1：单拍量预清零（锁存量 _eCause/_bFault/_bLeakNg/_fPrStart/_bBusyPrev 不入清单，R107） —— *)
_bDone    := FALSE;                                                                             // 完成脉冲预清 / Completion pulse preset
_bAborted := FALSE;                                                                             // 中止脉冲预清 / Abort pulse preset
bError    := FALSE;                                                                             // 故障标志预清（R45 配对） / Error preset
_bVent    := FALSE;                                                                             // 放气阀内部位预清（每拍显式赋值，R285） / Vent bit preset
fLeakRateKpaPerS := 0.0;                                                                        // 漏率出口预置 / Leak-rate outlet preset
_fRate    := 0.0;                                                                               // 速率工作值预置 / Rate working value preset

(* —— 段 2：组态闸（非法即锁存） —— *)
IF _bCfgBad THEN
    _eCause := E_DL_CpdCause.eCfgIllegal;                                                       // 归因：组态非法 / Cause: illegal configuration
    _bFault := TRUE;                                                                            // 锁存 / Latch
    _eState := E_DL_CpdPhase.eFault;                                                            // 入故障相 / Enter fault phase
END_IF

(* —— 段 3：迁出链（bReset 上升沿 → 待机相；清漏率锁存） —— *)
IF rtReset.Q THEN
    _bFault  := FALSE;                                                                          // 清故障锁存 / Clear fault latch
    _bLeakNg := FALSE;                                                                          // 清漏率锁存 / Clear the leak latch
    _eCause  := E_DL_CpdCause.eNone;                                                            // 清成因 / Clear cause
    _nWinCnt := 0;                                                                              // 窗计数清零 / Window count cleared
    _eState  := E_DL_CpdPhase.eIdle;                                                            // 回待机相 / Back to idle
END_IF

(* —— 段 4：相迁移（顺控 + 漏率判据 + 放气限速） —— *)
IF (NOT _bFault) AND (NOT _bCfgBad) THEN
    _bPrOk := NOT ((fPrMeasKpa <> fPrMeasKpa) OR ((fPrMeasKpa - fPrMeasKpa) <> (fPrMeasKpa - fPrMeasKpa)));   // 压力样本有限性
    _fPrNow := fPrMeasKpa;                                                                       // 当拍压力工作值 / Pressure working value

    IF bStop AND (_eState <> E_DL_CpdPhase.eIdle) THEN
        _bAborted := TRUE;                                                                       // 中止脉冲 / Abort pulse
        _eState := E_DL_CpdPhase.eIdle;                                                          // 回待机相（出口侧泵/阀随相切断） / Back to idle
    ELSE
        CASE _eState OF

        E_DL_CpdPhase.eIdle:
            _nWinCnt := 0;                                                                       // 待机相清零窗计数 / Clear the window count in idle
            IF rtStart.Q THEN
                _eState := E_DL_CpdPhase.ePump;                                                  // 启动沿进抽气相 / Enter pumping
            END_IF

        E_DL_CpdPhase.ePump:
            IF _bPrOk AND (_fPrNow <= fPrTargetKpa) THEN
                _eState := E_DL_CpdPhase.eStab;                                                  // 达目标真空：进稳压相 / Target reached, stabilise
            ELSIF tonPumpTo.Q THEN
                _eCause := E_DL_CpdCause.ePumpTimeout;                                           // 归因：抽气超时 / Cause: pump timeout
                _bFault := TRUE;                                                                 // 锁存 / Latch
                _eState := E_DL_CpdPhase.eFault;                                                 // 入故障相 / Enter fault phase
            END_IF

        E_DL_CpdPhase.eStab:
            IF tonStabTo.Q THEN
                _fPrStart := _fPrNow;                                                            // 记录窗起压（稳压结束点） / Record the window-start pressure
                _nWinCnt  := 0;                                                                  // 窗计数清零 / Clear the window count
                _eState   := E_DL_CpdPhase.eLeak;                                                // 进复测相 / Enter the leak phase
            END_IF

        E_DL_CpdPhase.eLeak:
            IF _bPrOk THEN
                _nWinCnt := _nWinCnt + 1;                                                        // 窗内采样计数 +1 / Count this sample
            END_IF
            IF tonLeakWin.Q THEN
                _fDtS := UDINT_TO_LREAL(_nWinCnt) * fSampleS;                                    // 实际时长 = 计数 × 周期 / Effective duration
                IF (_nWinCnt < 1) OR (fSampleS <= 0.0) THEN
                    _eCause := E_DL_CpdCause.eCfgIllegal;                                        // 分母闸：无有效样本，判据不成立 / Denominator gate
                    _bFault := TRUE;                                                             // 锁存 / Latch
                    _eState := E_DL_CpdPhase.eFault;                                             // 入故障相 / Enter fault phase
                ELSE
                    _fRate := ABS(_fPrNow - _fPrStart) / _fDtS;                                   // 漏率 = |Δp| / Δt（绝对值口径） / Leak rate
                    fLeakRateKpaPerS := _fRate;                                                   // 漏率出口 / Leak-rate outlet
                    IF _fRate > fLeakMaxKpaPerS THEN
                        _bLeakNg := TRUE;                                                         // 漏率超限：锁存 / Leak beyond the limit: latch
                        _eCause := E_DL_CpdCause.eLeakNg;                                         // 归因：漏率超限 / Cause: leak NG
                        _bFault := TRUE;                                                          // 故障锁存 / Latch the fault
                        _eState := E_DL_CpdPhase.eFault;                                          // 入故障相（禁止放气，等人工） / Enter fault phase
                    ELSE
                        _fPrPrev := _fPrNow;                                                      // 记录放气基准压力 / Record the vent reference pressure
                        _eState := E_DL_CpdPhase.eVent;                                           // 漏率合格：进放气相 / Leak OK, enter venting
                    END_IF
                END_IF
            END_IF

        E_DL_CpdPhase.eVent:
            IF _bPrOk THEN
                _fDtS  := fSampleS;                                                              // 单拍时长即采样周期（已过正域闸） / One-scan duration equals the sampling period
                _fRate := ABS(_fPrNow - _fPrPrev) / _fDtS;                                        // 逐拍放气速率 / Per-scan vent rate
                IF _fRate > fVentRateMaxKpaPerS THEN
                    _bVent := FALSE;                                                              // 超速：当拍关阀（占空比限速） / Too fast: close this scan
                    _eCause := E_DL_CpdCause.eVentTooFast;                                        // 归因：放气超速（信息级，不锁存） / Cause: vent too fast, info level
                ELSE
                    _bVent := TRUE;                                                               // 未超速：保持放气 / Below the limit: keep venting
                END_IF
                _fPrPrev := _fPrNow;                                                              // 更新基准压力 / Update the reference
            END_IF
            IF _bPrOk AND (_fPrNow >= 0.0) THEN
                _eState := E_DL_CpdPhase.eIdle;                                                  // 到常压：回待机相 / Atmosphere reached, back to idle
            ELSIF tonVentTo.Q THEN
                _eCause := E_DL_CpdCause.eVentTimeout;                                            // 归因：放气超时 / Cause: vent timeout
                _bFault := TRUE;                                                                  // 锁存 / Latch
                _eState := E_DL_CpdPhase.eFault;                                                  // 入故障相 / Enter fault phase
            END_IF

        E_DL_CpdPhase.eFault:
            ;                                                                                    // 故障相：仅等复位沿 / Wait for the reset edge only

        ELSE
            _eCause := E_DL_CpdCause.ePhaseBad;                                                  // 归因：非法相位 / Cause: illegal phase
            _bFault := TRUE;                                                                     // 锁存 / Latch
            _eState := E_DL_CpdPhase.eFault;                                                     // 强拉故障相 / Force fault phase

        END_CASE
    END_IF
END_IF

(* —— 段 5：完成脉冲（忙碌 → 待机，且无中止无故障；两段式单拍） —— *)
IF _bBusyPrev AND (_eState = E_DL_CpdPhase.eIdle) AND (NOT _bAborted) AND (NOT _bFault) THEN
    _bDone := TRUE;                                                                              // 完成脉冲 / Completion pulse
END_IF
_bBusyPrev := (_eState <> E_DL_CpdPhase.eIdle) AND (_eState <> E_DL_CpdPhase.eFault);            // 忙碌快照（本拍末） / Busy snapshot at body end

(* —— 段 6：出口单点映射（泵阀随相切断，名实双出口，R191） —— *)
bPumpValve := (_eState = E_DL_CpdPhase.ePump) OR (_eState = E_DL_CpdPhase.eStab) OR (_eState = E_DL_CpdPhase.eLeak);   // 抽气阀在前三相保持
bBusy      := (_eState <> E_DL_CpdPhase.eIdle) AND (_eState <> E_DL_CpdPhase.eFault);            // 忙碌 / Busy
bDone      := _bDone;                                                                            // 完成脉冲出口 / Completion pulse outlet
bAborted   := _bAborted;                                                                         // 中止脉冲出口 / Abort pulse outlet
bVentValve := _bVent AND (_eState = E_DL_CpdPhase.eVent);                                        // 放气阀位（仅放气相，单点映射） / Vent valve, vent phase only
bLeakNg    := _bLeakNg;                                                                          // 漏率锁存出口 / Leak latch outlet
ePhase     := _eState;                                                                           // 相出口 / Phase outlet
eCause     := _eCause;                                                                           // 成因出口 / Cause outlet
bError     := _bFault;                                                                           // 故障标志 / Error flag

END_FUNCTION_BLOCK

(* ---- FB_DL_ChuckVacuumSeq.st ---- *)
(*==============================================================================
 * 组件名称 (Component)  : FB_DL_ChuckVacuumSeq
 * 所属子库 (Sublibrary) : DL_Process
 * 当前版本 (Version)    : 1.0.0
 * 兼容性   (Platform)   : CODESYS 3.5+ / TwinCAT 3 / 汇川 InoProShop / 施耐德 Machine Expert
 *                         仅依赖 Standard.library（TON / R_TRIG），零厂商私有库
 * 功能描述 (Function)   : 卡盘真空吸附 / 释放顺控（四段：吸附 → 到位确认 → 加工互锁 → 破空释放）。
 *                         每相一枚**专用** TON，PT 各绑一个时间引脚，绝不共用实例改 PT：
 *                           eVacOn   吸附  ：tonVacTo  PT = tVacTo   （到位 bVacOk 即过相）
 *                           eConfirm 确认  ：tonConfTo PT = tConfirm （纯定时确认窗，窗内真空须保持）
 *                           eClamp   加工  ：无计时器，等 bProcessDone（外部加工完成）
 *                           eVent    释放  ：tonVentTo PT = tVentTo  （到位 bVentOk 即回待机）
 *                         到位判据：吸附相"定时到但未到位" → eVacTimeout；释放相"定时到但未破空" →
 *                         eVentTimeout；确认窗内真空掉落 → eVacLost（真空夹持不可中断）。
 *                         **加工互锁先于顺控**：加工进行中（bProcessActive）拒绝释放请求
 *                         （bReleaseReq），只置 bReleaseBlocked 单拍，不改变相（互锁优先级最高）。
 *                         验收向量：
 *                           ① 启动 → bVacValve 开；bVacOk 到 → eConfirm；tConfirm 到 → eClamp
 *                           ② eClamp 且 bProcessActive 时按释放请求 → 拒绝（bReleaseBlocked 单拍）
 *                           ③ bProcessDone 到 → eVent：bVacValve 关、bVentValve 开；bVentOk 到 → eIdle
 *                           ④ eVacOn 超时未到位 → eVacTimeout 锁存；eConfirm 窗内真空掉 → eVacLost 锁存
 * 接口     (Interface)  : 入 bStart 启动沿、bVacOk 真空到位、bVentOk 破空到位、bProcessDone 加工完成、
 *                         bProcessActive 加工进行中（互锁源）、bReleaseReq 释放请求、bStop 中止、
 *                         tVacTo 吸附超时、tConfirm 确认窗、tVentTo 破空超时、bReset 复位沿；
 *                         出 bVacValve 真空阀位、bVentValve 破空阀位、bClamped 夹持中、
 *                         bBusy 顺控进行中、bDone 完成脉冲（单拍）、bAborted 中止脉冲（单拍）、
 *                         bReleaseBlocked 释放被互锁拒绝（单拍）、ePhase 当前相、eCause 成因、bError 故障标志。
 * 边界     (Boundary)   : ① **属主边界（写死）：本件只出阀位与夹持指示，不驱动真空发生器/
 *                         电磁阀线圈、不判晶圆是否在位**（属 IO 映射层与在位检测件）；
 *                         ② **组态闸**：三个时间 ≤ T#0S → 锁存 eCfgIllegal；**互锁一致性闸**：
 *                         bProcessActive 为真而本件处于释放相 → 锁存 eInterlockViolation（防止外部
 *                         互锁源与顺控相位脱节）；
 *                         ③ **一相一 TON**：三枚专用 TON 在段 0 无条件调用，IN 由"当前相"表达式派生，
 *                         进相计时、出相复位，无跨相累积（R228A/R275）；
 *                         ④ **相驻留失守**：eConfirm 相真空掉落 → 立即落故障（驻留条件失守，R163）；
 *                         ⑤ **eFault 可迁出**：bReset 上升沿 → eIdle；bStop 亦可在非故障相回 eIdle，
 *                         但 eClamp 相中止需先破空，故中止统一走 eVent 相（安全侧）；
 *                         ⑥ 零全局耦合、零物理地址。
 * 分工声明 (Scope)      : 本件只管"卡盘吸附/释放四段时序与加工互锁"。不接管：真空度模拟量判读
 *                         （属模拟量件）、吸盘环真空（属 FB_DL_VacCupRingCtrl）、
 *                         腔体抽真空（属 FB_DL_ChamberPumpDownSeq）。
 * 来源标签 (Source Tag) : ROADMAP 空勾真缺口 P1（卡盘真空序，自研 clean-room）
 * 码表     (Codes)      : 本件不占用任何全局数字码位（零码位范式 R297）；诊断由 BOOL + ENUM 出口承担。
 * 红线自检 (Redline)    : R1 ✓ 零 GVL/VAR_EXTERNAL ｜ R2 ✓ 零 %I/%Q/%M ｜ R3 ✓ 纯 IEC 61131-3
 *                         R4 ✓ 组态闸 + 相超时 + 互锁一致性闸 + 驻留失守 ｜ R5 ✓ 声明逐行同行双语注释
 *                         R6 ✓ ENUM+CASE 含 ELSE 兜底 ｜ R7 ✓ 三 TON/两 R_TRIG 段 0 无条件刷新
 * 修订历史 (Revision)   : 2026-11-19  v1.0.0  R47 首版（批次 3 · 序号 13）
 *==============================================================================*)

TYPE E_DL_CvsPhase :
(
    eIdle   := 0,    // 待机相（阀位全关） / Idle, valves closed
    eVacOn  := 10,   // 吸附相（抽真空等到位） / Vacuum-on, waiting for vacuum
    eConfirm:= 20,   // 确认相（真空保持确认窗） / Confirmation window
    eClamp  := 30,   // 加工相（夹持中，等加工完成） / Clamped, waiting for process completion
    eVent   := 40,   // 释放相（破空等到位） / Venting, waiting for atmosphere
    eFault  := 90    // 故障相（等复位） / Fault, awaiting reset
);
END_TYPE

TYPE E_DL_CvsCause :
(
    eNone            := 0,   // 无异常 / No anomaly
    eCfgIllegal      := 1,   // 组态非法（时间非正） / Illegal configuration
    eVacTimeout      := 2,   // 吸附超时未到位 / Vacuum timeout
    eVentTimeout     := 3,   // 破空超时未到位 / Vent timeout
    eVacLost         := 4,   // 确认窗内真空掉（驻留失守） / Vacuum lost inside the confirmation window
    eInterlockViolation:= 5, // 互锁相位矛盾（加工中处于释放相） / Interlock contradiction
    ePhaseBad        := 6    // 非法相位兜底 / Illegal phase fallback
);
END_TYPE

FUNCTION_BLOCK FB_DL_ChuckVacuumSeq
VAR_INPUT
    bStart         : BOOL := FALSE;   // 启动沿，进入吸附相 [-] / Start edge, enters vacuum-on
    bVacOk         : BOOL := FALSE;   // 真空到位信号 [-] / Vacuum reached
    bVentOk        : BOOL := FALSE;   // 破空到位信号 [-] / Atmosphere reached
    bProcessDone   : BOOL := FALSE;   // 加工完成信号 [-] / Process finished
    bProcessActive : BOOL := FALSE;   // 加工进行中（互锁源，TRUE 时禁释放） [-] / Process active, release inhibited
    bReleaseReq    : BOOL := FALSE;   // 释放请求 [-] / Release request
    bStop          : BOOL := FALSE;   // 中止（安全侧：先进破空再回待机） [-] / Abort, vents first
    tVacTo         : TIME := T#10S;   // 吸附超时，域 > T#0S [ms] / Vacuum timeout
    tConfirm       : TIME := T#2S;    // 真空保持确认窗，域 > T#0S [ms] / Vacuum-hold confirmation window
    tVentTo        : TIME := T#10S;   // 破空超时，域 > T#0S [ms] / Vent timeout
    bReset         : BOOL := FALSE;   // 故障复位沿 [-] / Fault reset edge
END_VAR
VAR_OUTPUT
    bVacValve   : BOOL := FALSE;                          // 真空阀位 [-] / Vacuum valve position
    bVentValve  : BOOL := FALSE;                          // 破空阀位 [-] / Vent valve position
    bClamped    : BOOL := FALSE;                          // 夹持中（真空建立且确认过） [-] / Clamped
    bBusy       : BOOL := FALSE;                          // 顺控进行中 [-] / Sequence busy
    bDone       : BOOL := FALSE;                          // 完成脉冲（单拍） [-] / Completion pulse, single scan
    bAborted    : BOOL := FALSE;                          // 中止脉冲（单拍） [-] / Abort pulse, single scan
    bReleaseBlocked : BOOL := FALSE;                      // 释放被互锁拒绝（单拍） [-] / Release blocked by the interlock
    ePhase      : E_DL_CvsPhase := E_DL_CvsPhase.eIdle;   // 当前相出口 [-] / Present phase outlet
    eCause      : E_DL_CvsCause := E_DL_CvsCause.eNone;   // 成因出口（R190 归因唯一） [-] / Cause outlet
    bError      : BOOL := FALSE;                          // 故障标志 [-] / Error flag
END_VAR
VAR
    _eState    : E_DL_CvsPhase := E_DL_CvsPhase.eIdle;    // 内部相（CASE 唯一写入目标） / Internal phase
    _eCause    : E_DL_CvsCause := E_DL_CvsCause.eNone;    // 成因锁存量 / Latched cause
    _bFault    : BOOL := FALSE;                           // 故障锁存位 / Latched fault bit
    _bDone     : BOOL := FALSE;                           // 完成脉冲内部位（单拍） / Internal completion pulse
    _bAborted  : BOOL := FALSE;                           // 中止脉冲内部位（单拍） / Internal abort pulse
    _bRelBlock : BOOL := FALSE;                           // 释放被拒内部位（单拍） / Internal release-blocked flag
    _bCfgBad   : BOOL := FALSE;                           // 组态非法当拍量 / Illegal configuration this scan
    _bBusyPrev : BOOL := FALSE;                           // 上拍忙碌快照 / Busy snapshot of the previous scan
    tonVacTo   : TON;                                     // 吸附相专用超时，段 0 无条件调用 / Vacuum dedicated timeout
    tonConfTo  : TON;                                     // 确认相专用窗，段 0 无条件调用 / Confirmation dedicated window
    tonVentTo  : TON;                                     // 释放相专用超时，段 0 无条件调用 / Vent dedicated timeout
    rtStart    : R_TRIG;                                  // 启动沿实例，段 0 无条件调用 / Start edge instance
    rtReset    : R_TRIG;                                  // 复位沿实例，段 0 无条件调用 / Reset edge instance
END_VAR
VAR CONSTANT
    DL_CVS_MS   : INT := 0;               // 占位性零值常量（保持常量区非空，非事件码） [-] / Zero constant, not an event code
END_VAR

(* —— 段 0：组态闸 + 三枚专用 TON 与两沿无条件周期刷新（R228A/R275） —— *)
_bCfgBad := (tVacTo <= T#0S) OR (tConfirm <= T#0S) OR (tVentTo <= T#0S);                    // 三时间须为正 / All three times positive
rtStart(CLK := bStart);                                                                      // 启动沿 / Start edge
rtReset(CLK := bReset);                                                                      // 复位沿 / Reset edge
tonVacTo(IN := (_eState = E_DL_CvsPhase.eVacOn), PT := tVacTo);                               // 吸附相专用超时 / Vacuum timeout
tonConfTo(IN := (_eState = E_DL_CvsPhase.eConfirm), PT := tConfirm);                          // 确认相专用窗 / Confirmation window
tonVentTo(IN := (_eState = E_DL_CvsPhase.eVent), PT := tVentTo);                              // 释放相专用超时 / Vent timeout

(* —— 段 1：单拍量预清零（锁存量 _eCause/_bFault/_bBusyPrev 不入清单，R107） —— *)
_bDone     := FALSE;                                                                          // 完成脉冲预清 / Completion pulse preset
_bAborted  := FALSE;                                                                          // 中止脉冲预清 / Abort pulse preset
_bRelBlock := FALSE;                                                                          // 释放被拒预清 / Release-blocked preset
bError     := FALSE;                                                                          // 故障标志预清（R45 配对） / Error preset

(* —— 段 2：组态闸（时间非正即锁存） —— *)
IF _bCfgBad THEN
    _eCause := E_DL_CvsCause.eCfgIllegal;                                                    // 归因：组态非法 / Cause: illegal configuration
    _bFault := TRUE;                                                                          // 锁存 / Latch
    _eState := E_DL_CvsPhase.eFault;                                                          // 入故障相 / Enter fault phase
END_IF

(* —— 段 3：迁出链（bReset 上升沿 → 待机相；解除式恒可达） —— *)
IF rtReset.Q THEN
    _bFault := FALSE;                                                                          // 清故障锁存 / Clear fault latch
    _eCause := E_DL_CvsCause.eNone;                                                            // 清成因 / Clear cause
    _eState := E_DL_CvsPhase.eIdle;                                                            // 回待机相 / Back to idle
END_IF

(* —— 段 4：相迁移（顺控 + 互锁；互锁判定先于顺控推进） —— *)
IF (NOT _bFault) AND (NOT _bCfgBad) THEN
    CASE _eState OF

    E_DL_CvsPhase.eIdle:
        IF rtStart.Q THEN
            _eState := E_DL_CvsPhase.eVacOn;                                                   // 启动沿进吸附相 / Enter vacuum-on
        END_IF

    E_DL_CvsPhase.eVacOn:
        IF bVacOk THEN
            _eState := E_DL_CvsPhase.eConfirm;                                                 // 到位：进确认相 / Vacuum reached, enter confirmation
        ELSIF tonVacTo.Q THEN
            _eCause := E_DL_CvsCause.eVacTimeout;                                              // 归因：吸附超时 / Cause: vacuum timeout
            _bFault := TRUE;                                                                   // 锁存 / Latch
            _eState := E_DL_CvsPhase.eFault;                                                   // 入故障相 / Enter fault phase
        ELSIF bStop THEN
            _bAborted := TRUE;                                                                 // 中止脉冲 / Abort pulse
            _eState := E_DL_CvsPhase.eVent;                                                     // 中止先进破空（安全侧） / Abort vents first
        END_IF

    E_DL_CvsPhase.eConfirm:
        IF NOT bVacOk THEN
            _eCause := E_DL_CvsCause.eVacLost;                                                 // 驻留失守：确认窗内真空掉 / Vacuum lost, residency breach
            _bFault := TRUE;                                                                   // 锁存 / Latch
            _eState := E_DL_CvsPhase.eFault;                                                   // 入故障相 / Enter fault phase
        ELSIF tonConfTo.Q THEN
            _eState := E_DL_CvsPhase.eClamp;                                                    // 确认窗满：进加工相 / Confirmed, enter the clamp phase
        END_IF

    E_DL_CvsPhase.eClamp:
        IF bReleaseReq AND bProcessActive THEN
            _bRelBlock := TRUE;                                                                // 加工中拒释放（互锁先于顺控） / Release blocked while processing
        ELSIF (bReleaseReq AND bProcessDone) OR bStop THEN
            _bAborted := bStop AND (NOT bProcessDone);                                          // 中止（无完成）置中止脉冲 / Abort pulse only on stop
            _eState := E_DL_CvsPhase.eVent;                                                     // 进破空相 / Enter venting
        END_IF

    E_DL_CvsPhase.eVent:
        IF bVentOk THEN
            _eState := E_DL_CvsPhase.eIdle;                                                     // 破空到位：回待机相 / Atmosphere reached, back to idle
        ELSIF tonVentTo.Q THEN
            _eCause := E_DL_CvsCause.eVentTimeout;                                              // 归因：破空超时 / Cause: vent timeout
            _bFault := TRUE;                                                                   // 锁存 / Latch
            _eState := E_DL_CvsPhase.eFault;                                                   // 入故障相 / Enter fault phase
        END_IF

    E_DL_CvsPhase.eFault:
        ;                                                                                      // 故障相：仅等复位沿 / Wait for the reset edge only

    ELSE
        _eCause := E_DL_CvsCause.ePhaseBad;                                                    // 归因：非法相位 / Cause: illegal phase
        _bFault := TRUE;                                                                       // 锁存 / Latch
        _eState := E_DL_CvsPhase.eFault;                                                       // 强拉故障相 / Force fault phase

    END_CASE
END_IF

(* —— 段 5：互锁一致性闸（加工中却处于释放/待机相 → 相位与外部互锁源脱节） —— *)
IF bProcessActive AND ((_eState = E_DL_CvsPhase.eVent) OR (_eState = E_DL_CvsPhase.eIdle)) THEN
    _eCause := E_DL_CvsCause.eInterlockViolation;                                              // 归因：互锁相位矛盾 / Cause: interlock contradiction
    _bFault := TRUE;                                                                            // 锁存 / Latch
    _eState := E_DL_CvsPhase.eFault;                                                            // 入故障相 / Enter fault phase
END_IF

(* —— 段 6：完成脉冲（忙碌 → 待机且无中止无故障；两段式单拍） —— *)
IF _bBusyPrev AND (_eState = E_DL_CvsPhase.eIdle) AND (NOT _bAborted) AND (NOT _bFault) THEN
    _bDone := TRUE;                                                                             // 完成脉冲 / Completion pulse
END_IF
_bBusyPrev := (_eState <> E_DL_CvsPhase.eIdle) AND (_eState <> E_DL_CvsPhase.eFault);           // 忙碌快照（本拍末） / Busy snapshot at body end

(* —— 段 7：出口单点映射（阀位与相/夹持同源，R191） —— *)
bVacValve  := ((_eState = E_DL_CvsPhase.eVacOn) OR (_eState = E_DL_CvsPhase.eConfirm) OR (_eState = E_DL_CvsPhase.eClamp))
              AND (NOT _bFault);                                                                // 吸附/确认/加工相保持真空（故障相切断） / Vacuum held in three phases only
bVentValve := (_eState = E_DL_CvsPhase.eVent);                                                  // 破空阀仅在释放相 / Vent valve only in the vent phase
bClamped   := (_eState = E_DL_CvsPhase.eClamp);                                                 // 夹持指示 / Clamped indicator
bBusy      := (_eState <> E_DL_CvsPhase.eIdle) AND (_eState <> E_DL_CvsPhase.eFault);           // 忙碌 / Busy
bDone      := _bDone;                                                                           // 完成脉冲出口 / Completion pulse outlet
bAborted   := _bAborted;                                                                        // 中止脉冲出口 / Abort pulse outlet
bReleaseBlocked := _bRelBlock;                                                                  // 释放被拒出口 / Release-blocked outlet
ePhase     := _eState;                                                                          // 相出口 / Phase outlet
eCause     := _eCause;                                                                          // 成因出口 / Cause outlet
bError     := _bFault;                                                                          // 故障标志 / Error flag

END_FUNCTION_BLOCK
